RESOURCE RES0 : EMB_RES_ECO
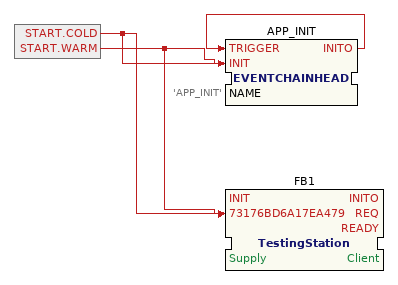
  FBS
    FB1 : TestingStation;
    APP_INIT : EVENTCHAINHEAD(NAME := 'APP_INIT');
  END_FBS
  EVENT_CONNECTIONS
    APP_INIT.INITO TO APP_INIT.TRIGGER;
    START.COLD TO APP_INIT.INIT;
    START.WARM TO APP_INIT.INIT;
    START.COLD TO FB1.73176BD6A17EA479;
    START.WARM TO FB1.73176BD6A17EA479;
  END_CONNECTIONS
END_RESOURCE
